FUNCTION_BLOCK BtnController (* Basic Function Block Type *)
  (* Standard: 61499-2 *)
  (* Version 0.0, 10/20/2026, macie, Schneider Electric, Template *)
  PACKAGE Main;
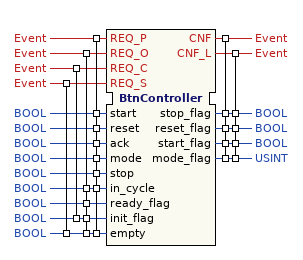
  EVENT_INPUT
    REQ_P WITH start, reset, ack, mode, stop, in_cycle, empty; (* Normal Execution Request *)
    REQ_O WITH in_cycle, ready_flag, init_flag, empty;
    REQ_C WITH init_flag;
    REQ_S WITH empty;
  END_EVENT
  EVENT_OUTPUT
    CNF WITH stop_flag, reset_flag, start_flag, mode_flag; (* Execution Confirmation *)
    CNF_L WITH stop_flag, reset_flag, start_flag, mode_flag;
  END_EVENT
  VAR_INPUT
    start : BOOL; (* Input event qualifier *)
    reset : BOOL;
    ack : BOOL;
    mode : BOOL := TRUE;
    stop : BOOL;
    in_cycle : BOOL := FALSE;
    ready_flag : BOOL := TRUE;
    init_flag : BOOL;
    empty : BOOL;
  END_VAR
  VAR_OUTPUT
    stop_flag : BOOL := FALSE; (* Output event qualifier *)
    reset_flag : BOOL;
    start_flag : BOOL;
    mode_flag : USINT := 0;
  END_VAR
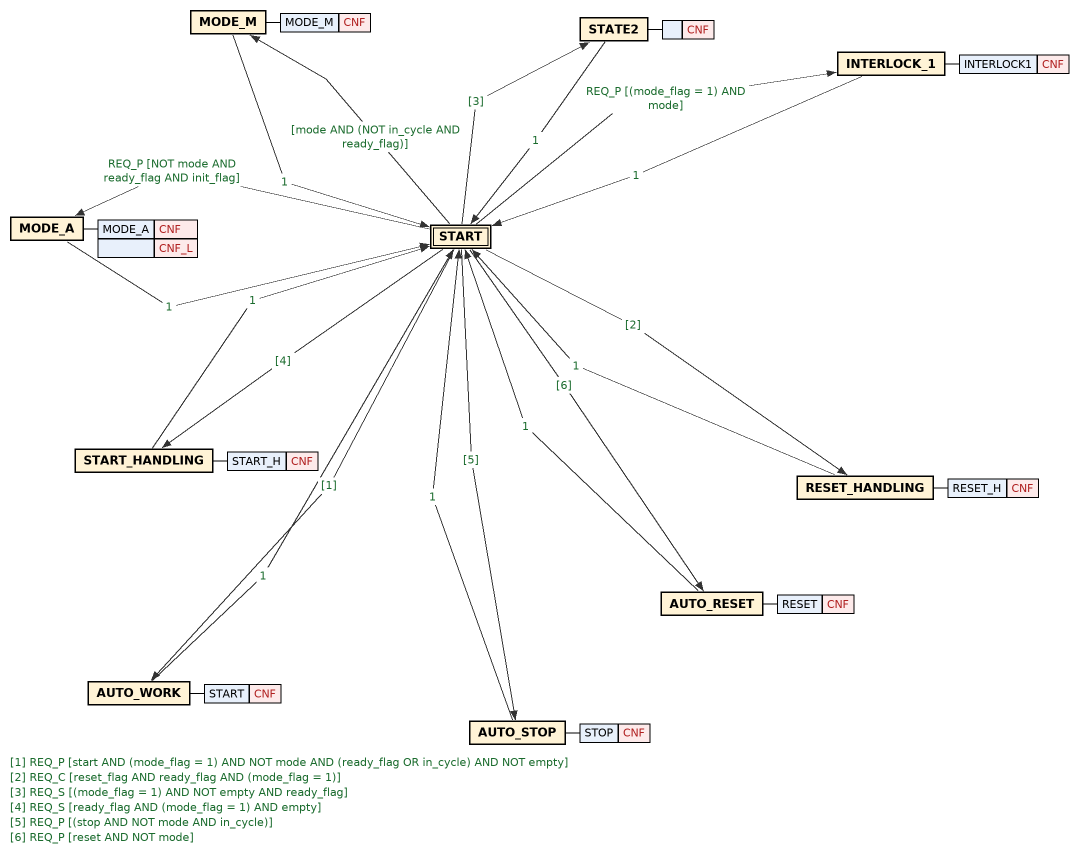
  EC_STATES
    START; (* Initial State *)
    AUTO_WORK : START -> CNF; (* Normal execution *)
    AUTO_STOP : STOP -> CNF;
    AUTO_RESET : RESET -> CNF;
    MODE_M : MODE_M -> CNF;
    MODE_A : MODE_A -> CNF, -> CNF_L;
    RESET_HANDLING : RESET_H -> CNF;
    STATE2 : -> CNF;
    START_HANDLING : START_H -> CNF;
    INTERLOCK_1 : INTERLOCK1 -> CNF;
  END_STATES
  EC_TRANSITIONS
    START TO AUTO_WORK := REQ_P [start AND (mode_flag = 1) AND NOT mode AND (ready_flag OR in_cycle) AND NOT empty];
    AUTO_WORK TO START := 1;
    START TO AUTO_STOP := REQ_P [(stop AND NOT mode AND in_cycle)];
    START TO AUTO_RESET := REQ_P [reset AND NOT mode];
    AUTO_RESET TO START := 1;
    AUTO_STOP TO START := 1;
    START TO MODE_M := [mode AND (NOT in_cycle AND ready_flag)];
    MODE_M TO START := 1;
    START TO MODE_A := REQ_P [NOT mode AND ready_flag AND init_flag];
    MODE_A TO START := 1;
    START TO RESET_HANDLING := REQ_C [reset_flag AND ready_flag AND (mode_flag = 1)];
    RESET_HANDLING TO START := 1;
    START TO STATE2 := REQ_S [(mode_flag = 1) AND NOT empty AND ready_flag];
    STATE2 TO START := 1;
    START TO START_HANDLING := REQ_S [ready_flag AND (mode_flag = 1) AND empty];
    START_HANDLING TO START := 1;
    START TO INTERLOCK_1 := REQ_P [(mode_flag = 1) AND mode];
    INTERLOCK_1 TO START := 1;
  END_TRANSITIONS
  ALGORITHM INIT IN ST: (* Initialization algorithm *)
;
  END_ALGORITHM
  ALGORITHM REQ IN ST: (* Normally executed algorithm *)
;
  END_ALGORITHM
  ALGORITHM START IN ST:
;
reset_flag := FALSE;
stop_flag := FALSE;
start_flag := TRUE;
  END_ALGORITHM
  ALGORITHM STOP IN ST:
;
stop_flag := TRUE;
start_flag := FALSE;
  END_ALGORITHM
  ALGORITHM RESET IN ST:
;
reset_flag := TRUE;
start_flag := FALSE;
stop_flag := FALSE;
  END_ALGORITHM
  ALGORITHM MODE_M IN ST:
;
mode_flag := 0;
  END_ALGORITHM
  ALGORITHM MODE_A IN ST:
;
mode_flag := 1;
//stop_flag := TRUE;
  END_ALGORITHM
  ALGORITHM RESET_H IN ST:
;
reset_flag := FALSE;
  END_ALGORITHM
  ALGORITHM START_H IN ST:
;
start_flag := FALSE;
  END_ALGORITHM
  ALGORITHM INTERLOCK1 IN ST:
;
stop_flag := TRUE;
start_flag := FALSE;
  END_ALGORITHM
END_FUNCTION_BLOCK
